Fanuc KAREL source: kf00088.KL

-- PROVISIONAL review KL for V940-1; original PC SHA256 1777a99b50431928b63fbd4a5098a7bdb57e2f13b65bc54c55eb167c1f6cc59e
-- Incomplete behavior may be omitted. Consult companion uncertainty JSON. Do not deploy.
PROGRAM KF00088
%NOLOCKGROUP
BEGIN
  -- V9_ZERO_TABLE_METADATA_HINT layout=0002_ascii; no indexed target words; source/name/runtime held
  -- UNRESOLVED_PC offsets 5-28; opcodes 27,22,1C,31,4A
  -- UNRESOLVED_PC offsets 33-37; opcodes 7F
END KF00088
